Fanuc KAREL source: ka00065.KL

PROGRAM KA00065
%STACKSIZE=65535
%PRIORITY=65535
%NOLOCKGROUP
VAR
SRC : XYZWPR
DST : POSITION
BEGIN
SRC.X=1.0
-- UNSAFE_SOURCE_IR line 8: DST = convert_xyzwpr_to_position(SRC)
END KA00065
